// TIA Portal V20 export
// export: Created 2026-10-11T05:26:44.7307727Z, ExportSetting WithDefaults, DisplayName Totally Integrated Automation Portal, DisplayVersion V20, DisplayName TIA Portal Openness, DisplayVersion V20, DisplayName TIA Portal Teamcenter Gateway, DisplayVersion V20, DisplayName TIA Portal Version Control Interface, DisplayVersion V20, DisplayName SINAMICS Startdrive Advanced, DisplayVersion V20 SP1 Update 2, DisplayName SINAMICS Startdrive G110M, G120, G120C, G120D, G120P, G115D, DisplayVersion V20 SP1 Update 2, DisplayName SINAMICS Startdrive G130, G150, S120, S150, SINAMICS MV, G220, S200, S210, DisplayVersion V20 SP1 Update 2, DisplayName STEP 7 Professional, DisplayVersion V20, DisplayName STEP 7 Safety, DisplayVersion V20, DisplayName WinCC Basic/Comfort/Advanced, DisplayVersion V20, DisplayName WinCC Professional, DisplayVersion V20, DisplayName WinCC Unified, DisplayVersion V20
FUNCTION "FRK_HistoryEvent" : Void   // FC52, SCL
{ S7_Optimized_Access := 'TRUE' }
VERSION : 0.1
// Shared Unit routing: typed generated edges carry these owning predicates.
// stored: AutoNumber true, IsIECCheckEnabled false, SetENOAutomatically false, UDAEnableTagReadback false
   VAR_INPUT
      Reason : DInt;
      Description : WString;
      SourcePath : WString;
   END_VAR
   VAR_IN_OUT
      History : Array[1..16] of "ST_Diagnostic";
      Head : Int;
   END_VAR
   VAR_TEMP
      Stamp : DTL;
      ResultCode : Int;
   END_VAR
BEGIN

   IF #Head < 0 OR #Head >= 16 THEN
       #Head := 0;
   END_IF;
   #Head := #Head + 1;
   #History[#Head] := "FRK_UnitScratch".EmptyDiagnostic;
   #History[#Head].ReasonCode := #Reason;
   #History[#Head].Description := #Description;
   #History[#Head].SourcePath := #SourcePath;
   #History[#Head].Severity := 0;
   #History[#Head].Category := 2;
   #ResultCode := RD_SYS_T(OUT => #Stamp);
   IF #ResultCode = 0 THEN
       #History[#Head].Since := DTL_TO_LDT(#Stamp);
   END_IF;
END_FUNCTION
